// TIA Portal V21 export
// export: Created 2026-08-21T20:18:51.9495594Z, ExportSetting None, DisplayName Totally Integrated Automation Portal, DisplayVersion V21, DisplayName STEP 7 Professional, DisplayVersion V21, DisplayName STEP 7 Safety, DisplayVersion V21, DisplayName Tech WebApplication, DisplayVersion V21, DisplayName WinCC Basic/Comfort/Advanced, DisplayVersion V21, DisplayName WinCC Professional, DisplayVersion V21, DisplayName WinCC Unified, DisplayVersion V21
DATA_BLOCK "ProcedureParameters_DB"   // DB33
AUTHOR : Siemens AG
FAMILY : ServiceControl
VERSION : 1.0
// stored: InstanceOfName ProcedureParameters, InstanceOfType FB
"ProcedureParameters"
   // VAR
   //    MTPAnalog { S7_SetPoint := 'True'} : Array[0..2] of "UDT_MTP_AnaServParam";
   //    MTPDigital { S7_SetPoint := 'True'} : Array[0..0] of "UDT_MTP_DIntServParam";
   //    MTPBinary { S7_SetPoint := 'True'} : Array[0..0] of "UDT_MTP_BinServParam";
   //    MTPString { S7_SetPoint := 'True'} : Array[0..0] of "UDT_MTP_StringServParam";
   // END_VAR
BEGIN
   MTPAnalog[0..2].Sync := True;
   MTPAnalog[0].VExt := 25.0;
   MTPAnalog[1].VExt := 1000.0;
   MTPAnalog[2].VExt := 10.0;
   MTPAnalog[0].VOp := 25.0;
   MTPAnalog[1].VOp := 1000.0;
   MTPAnalog[2].VOp := 10.0;
   MTPAnalog[0].VInt := 25.0;
   MTPAnalog[1].VInt := 1000.0;
   MTPAnalog[2].VInt := 10.0;
   MTPAnalog[0].VReq := 25.0;
   MTPAnalog[1].VReq := 1000.0;
   MTPAnalog[2].VReq := 10.0;
   MTPAnalog[0].VOut := 25.0;
   MTPAnalog[1].VOut := 1000.0;
   MTPAnalog[2].VOut := 10.0;
   MTPAnalog[0].VSclMin := 0.0;
   MTPAnalog[1].VSclMin := 100.0;
   MTPAnalog[2].VSclMin := 0.0;
   MTPAnalog[0].VSclMax := 32.0;
   MTPAnalog[1].VSclMax := 3000.0;
   MTPAnalog[2].VSclMax := 300.0;
   MTPAnalog[0].VUnit := 1600;
   MTPAnalog[1].VUnit := 1038;
   MTPAnalog[2].VUnit := 1054;
   MTPAnalog[0].VMin := 0.0;
   MTPAnalog[1].VMin := 100.0;
   MTPAnalog[2].VMin := 5.0;
   MTPAnalog[0].VMax := 32.0;
   MTPAnalog[1].VMax := 3000.0;
   MTPAnalog[2].VMax := 300.0;
END_DATA_BLOCK
